// TIA Portal V21 export
// export: Created 2026-11-21T13:26:58.5467574Z, ExportSetting WithDefaults, DisplayName Totally Integrated Automation Portal, DisplayVersion V21, DisplayName STEP 7 Professional, DisplayVersion V21, DisplayName STEP 7 Safety, DisplayVersion V21, DisplayName Tech WebApplication, DisplayVersion V21, DisplayName WinCC Basic/Comfort/Advanced, DisplayVersion V21, DisplayName WinCC Unified, DisplayVersion V21
FUNCTION_BLOCK "Tank"   // FB1, SCL
TITLE = Behälter überwachen / Watch the tank / Surveiller le réservoir
{ S7_Optimized_Access := 'TRUE' }
VERSION : 0.1
// Meldet einen hohen und einen niedrigen Füllstand. / Reports a high and a low level. / Signale un niveau haut et un niveau bas.
// stored: AutoNumber true, IsIECCheckEnabled false, IsRetainMemResEnabled false, MemoryReserve 100, SetENOAutomatically false, UDAEnableTagReadback false
   VAR_INPUT
      level : Int;   // Füllstand in mm
      high : Bool;   // Grenzwert oben erreicht
      low : Bool;
      state : Int;   // Zustand, Index in die Textliste States
   END_VAR
   VAR
      highAlarm { S7_SetPoint := 'True'} : Program_Alarm;
      lowAlarm { S7_SetPoint := 'True'} : Program_Alarm;
   END_VAR
BEGIN

    #highAlarm(SIG := #high, SD_1 := #level);
    #lowAlarm(SIG := #low, SD_1 := #level, SD_2 := #state);
END_FUNCTION_BLOCK
